(* IEC 61131-3 sources: IRIS-Project/LASAL CONTROL SOFTWARE/LasalProject_2025_09_12/Network/Manual, 1 file *)

(* ---- ONE_Manual_Table.st ---- *)
#define OBJECTS_CONFIG

FUNCTION GLOBAL TAB ONE_Manual
-1$UINT, 0$UINT,
0$UINT, 0$UINT,

5$UDINT,
TO_UDINT(3284677247), "AutoManSelector", 0$UINT, 0$UINT, 1$UINT,
TO_UDINT(453563333), "Manual_Motor", 0$UINT, 0$UINT, 3$UINT,
TO_UDINT(1187451384), "Manual_MotorBT", 0$UINT, 0$UINT, 1$UINT,
TO_UDINT(2321534941), "ManualMotor_CBCM", 0$UINT, 0$UINT, 2$UINT,
TO_UDINT(2579655818), "ManualMotor_DB", 0$UINT, 0$UINT, 1$UINT,

_NO_ATTR, TO_UDINT(1134906152), "AUTOMANSELECTOR1",

_NO_ATTR, TO_UDINT(3551337390), "M1_CHARGE_SLIDER",
_NO_ATTR, TO_UDINT(3029375565), "M3_DISCHARGE_SLIDER",
_NO_ATTR, TO_UDINT(1249984746), "M6_LONGITUDINAL_AXIS",

_NO_ATTR, TO_UDINT(3611066561), "M7_TARGET_BLOCK",

_NO_ATTR, TO_UDINT(1011716386), "M2_CHARGE_BUFFER",
_NO_ATTR, TO_UDINT(3210558052), "M5_CENTRAL_MOVEMENT",

_NO_ATTR, TO_UDINT(2871226588), "M4_DISCHARGE_BUFFER",

//Internal connections
0$UDINT,
0$UDINT,
0$UDINT,
21$UDINT,
TO_UDINT(0), "toManualM1", TO_UDINT(1), "Enable",
TO_UDINT(0), "toManualM2", TO_UDINT(5), "Enable",
TO_UDINT(0), "toManualM3", TO_UDINT(2), "Enable",
TO_UDINT(0), "toManualM4", TO_UDINT(7), "Enable",
TO_UDINT(0), "toManualM5", TO_UDINT(6), "Enable",
TO_UDINT(0), "toManualM6", TO_UDINT(3), "Enable",
TO_UDINT(0), "toManualM7", TO_UDINT(4), "Enable",
TO_UDINT(0), "StopM1", TO_UDINT(1), "Stop",
TO_UDINT(0), "StopM2", TO_UDINT(5), "Stop",
TO_UDINT(0), "StopM3", TO_UDINT(2), "Stop",
TO_UDINT(0), "StopM4", TO_UDINT(7), "Stop",
TO_UDINT(0), "StopM5", TO_UDINT(6), "Stop",
TO_UDINT(0), "StopM6", TO_UDINT(3), "Stop",
TO_UDINT(0), "StopM7", TO_UDINT(4), "Stop",
TO_UDINT(0), "ResetM1", TO_UDINT(1), "S_Reset",
TO_UDINT(0), "ResetM2", TO_UDINT(5), "S_Reset",
TO_UDINT(0), "ResetM3", TO_UDINT(2), "S_Reset",
TO_UDINT(0), "ResetM4", TO_UDINT(7), "S_Reset",
TO_UDINT(0), "ResetM5", TO_UDINT(6), "S_Reset",
TO_UDINT(0), "ResetM6", TO_UDINT(3), "S_Reset",
TO_UDINT(0), "ResetM7", TO_UDINT(4), "S_Reset",

//Initialization values
0$UDINT,
1$UDINT,
TO_UDINT(1), "Comando_Motore", TO_UDINT(PASSIVE_LMCAXIS),//|Manual.M1_Charge_Slider.Comando_Motore;

//Symbolic initialization values
0$UDINT,
0$UDINT,

//Initialization of string values
0$UDINT,
0$UDINT,

//Configuration of tasks (RealTime, Cyclic, Background)
0$UDINT,
0$UDINT,

0$UDINT,
8$UDINT,
TO_UDINT(0), (100)$UDINT, 4194303$DINT, 	//AUTOMANSELECTOR1
TO_UDINT(1), (100)$UDINT, 4194303$DINT, 	//M1_CHARGE_SLIDER
TO_UDINT(2), (100)$UDINT, 4194303$DINT, 	//M3_DISCHARGE_SLIDER
TO_UDINT(3), (100)$UDINT, 4194303$DINT, 	//M6_LONGITUDINAL_AXIS
TO_UDINT(4), (100)$UDINT, 4194303$DINT, 	//M7_TARGET_BLOCK
TO_UDINT(5), (100)$UDINT, 4194303$DINT, 	//M2_CHARGE_BUFFER
TO_UDINT(6), (100)$UDINT, 4194303$DINT, 	//M5_CENTRAL_MOVEMENT
TO_UDINT(7), (100)$UDINT, 4194303$DINT, 	//M4_DISCHARGE_BUFFER

0$UDINT,
0$UDINT,

//External connections
0$UDINT,
34$UDINT,
TO_UDINT(0), "toAutomatic", C_DIR, TO_UDINT(1533940179), "Manager_globale1","enable",
TO_UDINT(0), "c_EasyGUIEn_MainS", C_DIR, TO_UDINT(3321030168), "MainSequence1","s_EasyGUI",
TO_UDINT(0), "c_EasyGUIEn_IrrT", C_DIR, TO_UDINT(101499717), "IrradiationTimers","s_EasyGUI",
TO_UDINT(1), "Comando_Motore", C_TRY, TO_UDINT(1906010274), "_LMCAxis_M1","Control",
TO_UDINT(1), "M_LS_1", C_TRY, TO_UDINT(201264582), "ST1511","Input1",
TO_UDINT(1), "M_LS_2", C_TRY, TO_UDINT(201264582), "ST1511","Input2",
TO_UDINT(1), "setPositionController", C_DIR, TO_UDINT(1906010274), "_LMCAxis_M1","ActPos",
TO_UDINT(1), "c_MaxCurrent", C_DIR, TO_UDINT(201264582), "ST1511","MaxCurrent",
TO_UDINT(2), "Comando_Motore", C_TRY, TO_UDINT(2677344654), "_LMCAxis_M3","Control",
TO_UDINT(2), "M_LS_1", C_TRY, TO_UDINT(3857804522), "ST1513","Input2",
TO_UDINT(2), "M_LS_2", C_TRY, TO_UDINT(3857804522), "ST1513","Input1",
TO_UDINT(2), "setPositionController", C_DIR, TO_UDINT(2677344654), "_LMCAxis_M3","ActPos",
TO_UDINT(2), "c_MaxCurrent", C_DIR, TO_UDINT(3857804522), "ST1513","MaxCurrent",
TO_UDINT(3), "Comando_Motore", C_TRY, TO_UDINT(4026531073), "_LMCAxis_M6","Control",
TO_UDINT(3), "M_LS_1", C_TRY, TO_UDINT(2510002277), "ST1516","Input1",
TO_UDINT(3), "M_LS_2", C_TRY, TO_UDINT(2510002277), "ST1516","Input2",
TO_UDINT(3), "setPositionController", C_DIR, TO_UDINT(4026531073), "_LMCAxis_M6","ActPos",
TO_UDINT(3), "c_MaxCurrent", C_DIR, TO_UDINT(2510002277), "ST1516","MaxCurrent",
TO_UDINT(4), "Comando_Motore", C_TRY, TO_UDINT(2566442391), "_LMCAxis_M7","Control",
TO_UDINT(4), "M_LS_1", C_TRY, TO_UDINT(3801917683), "ST1517","Input1",
TO_UDINT(4), "M_LS_2", C_TRY, TO_UDINT(3801917683), "ST1517","Input2",
TO_UDINT(4), "setPositionController", C_DIR, TO_UDINT(2566442391), "_LMCAxis_M7","ActPos",
TO_UDINT(5), "Comando_Motore", C_TRY, TO_UDINT(3901896984), "_LMCAxis_M2","Control",
TO_UDINT(5), "M_LS", C_TRY, TO_UDINT(2465619068), "ST1512","Input2",
TO_UDINT(5), "setPositionController", C_DIR, TO_UDINT(3901896984), "_LMCAxis_M2","ActPos",
TO_UDINT(5), "c_MaxCurrent", C_DIR, TO_UDINT(2465619068), "ST1512","MaxCurrent",
TO_UDINT(6), "Comando_Motore", C_TRY, TO_UDINT(1995877563), "_LMCAxis_M5","Control",
TO_UDINT(6), "M_LS", C_TRY, TO_UDINT(210946527), "ST1515","Input1",
TO_UDINT(6), "setPositionController", C_DIR, TO_UDINT(1995877563), "_LMCAxis_M5","ActPos",
TO_UDINT(6), "c_MaxCurrent", C_DIR, TO_UDINT(210946527), "ST1515","MaxCurrent",
TO_UDINT(7), "Comando_Motore", C_TRY, TO_UDINT(32611373), "_LMCAxis_M4","Control",
TO_UDINT(7), "M_LS", C_TRY, TO_UDINT(2073426249), "ST1514","Input1",
TO_UDINT(7), "setPositionController", C_DIR, TO_UDINT(32611373), "_LMCAxis_M4","ActPos",
TO_UDINT(7), "c_MaxCurrent", C_DIR, TO_UDINT(2073426249), "ST1514","MaxCurrent",

//Magic internal connections
0$UDINT,
0$UDINT,

//Configuration of timeslots of tasks (RealTime, Cyclic)
#ifdef __LSLLDR_TIMESLOTS__
0$UDINT,
0$UDINT,

0$UDINT,
0$UDINT,

#endif //__LSLLDR_TIMESLOTS__

//MultiMaster connections
#ifdef __LSLLDR_MULTIMASTER__
0$UDINT,
0$UDINT,
#endif //__LSLLDR_MULTIMASTER__

//Configuration for task ID (RealTime, CyclicTime)
#ifdef __LSLLDR_TASKID__
"\\\\TASKS2  "
0$UDINT,
0$UDINT,

0$UDINT,
8$UDINT,
(0)$UDINT, 	//AUTOMANSELECTOR1
(0)$UDINT, 	//M1_CHARGE_SLIDER
(0)$UDINT, 	//M3_DISCHARGE_SLIDER
(0)$UDINT, 	//M6_LONGITUDINAL_AXIS
(0)$UDINT, 	//M7_TARGET_BLOCK
(0)$UDINT, 	//M2_CHARGE_BUFFER
(0)$UDINT, 	//M5_CENTRAL_MOVEMENT
(0)$UDINT, 	//M4_DISCHARGE_BUFFER

0$UDINT,
0$UDINT,

#endif //__LSLLDR_TASKID__

END_FUNCTION
